(* PLC project probe, plc-portfolio cds2astra probe 0.1.0 *)
(* stored: creationDateTime 2026-10-20T00:00:00, modificationDateTime 2026-10-20T00:00:00 *)

PROGRAM PRG_P2
VAR
END_VAR

                    GVL_P2.iCount := GVL_P2.iCount + 1;
                  
END_PROGRAM

PROGRAM PRG_P2Slow
VAR
END_VAR

                    ;
                  
END_PROGRAM

CONFIGURATION CfgOther
  RESOURCE ResOther ON PLC
(* global variable list GVL_P2 *)
VAR_GLOBAL
    iCount : INT;
END_VAR
    TASK T_Fast(INTERVAL := T#20ms, PRIORITY := 3);
    TASK T_Slow(INTERVAL := T#500ms, PRIORITY := 20);
    PROGRAM PRG_P2 WITH T_Fast : PRG_P2;
    PROGRAM PRG_P2Slow WITH T_Slow : PRG_P2Slow;
  END_RESOURCE
END_CONFIGURATION
